TYPE "ST_S11RecoveryControl"
VERSION : 0.1
   STRUCT
      SchemaVersion : UInt := 1;
      Go : Bool;
   END_STRUCT;
END_TYPE
